Staubli VAL3: unbind.pgx

program unbind()
begin
  userPageUnbind("editProg","lst1","value")
  userPageUnbind("editProg","lst1","options")
end
